// TIA Portal V21 export
// export: Created 2026-10-23T20:43:22.5556805Z, ExportSetting WithDefaults, DisplayName Totally Integrated Automation Portal, DisplayVersion V21 Update 1, DisplayName SINAMICS Startdrive Advanced, DisplayVersion V21 HF2, DisplayName SINAMICS Startdrive G110M, G120, G120C, G120D, G120P, G115D, DisplayVersion V21 HF2, DisplayName SINAMICS Startdrive G130, G150, S120, S150, G200, G220, S200, S210, S220, Innomotics MVD, DisplayVersion V21 HF2, DisplayName STEP 7 Professional, DisplayVersion V21 Update 1, DisplayName STEP 7 Safety, DisplayVersion V21, DisplayName Tech WebApplication, DisplayVersion V21, DisplayName WinCC Basic/Comfort/Advanced, DisplayVersion V21 Update 1, DisplayName WinCC Unified, DisplayVersion V21 Update 1
FUNCTION "FC_AnaCaseReal" : Int   // FC14, SCL
TITLE = Analyzer: CASE without ELSE, REAL compared with =
{ S7_Optimized_Access := 'TRUE' }
VERSION : 0.1
// Rule C26i: the CASE has no ELSE, and a REAL is compared with =
// stored: AutoNumber true, IsIECCheckEnabled false, SetENOAutomatically false, UDAEnableTagReadback false
   VAR_INPUT
      Mode : Int;   // Mode
      Level : Real;   // Level
   END_VAR
   VAR_TEMP
      Code : Int;   // Result code
   END_VAR
BEGIN

       #Code := 0;
       CASE #Mode OF
           1:
               #Code := 10;
           2:
               #Code := 20;
       END_CASE;
       IF #Level = 1.5 THEN
           #Code := #Code + 1;
       END_IF;
       #FC_AnaCaseReal := #Code;
END_FUNCTION
